Fanuc KAREL source: kf00097.KL

-- PROVISIONAL review KL for V1013-1; original PC SHA256 61d1d2d0537b2f02508713676a499a9c69016aa3983c12c6525e9969e3959a7d
-- Incomplete behavior may be omitted. Consult companion uncertainty JSON. Do not deploy.
PROGRAM KF00097
%NOLOCKGROUP
BEGIN
  -- UNRESOLVED_PC offsets 5-16; opcodes 2E,23
  -- UNRESOLVED_PC offsets 21-32; opcodes 2E,23
  -- UNRESOLVED_PC offsets 37-55; opcodes 27,27,9D,22,22,31
  -- UNRESOLVED_PC offsets 60-64; opcodes 7F
END KF00097
